Fanuc KAREL source: kt00240.KL

PROGRAM KT00240
%STACKSIZE=65535
%PRIORITY=65535
%NOLOCKGROUP
VAR
I1 : INTEGER
H2 : ARRAY[2] OF SHORT
OUT : INTEGER
BEGIN
I1=2
H2[1]=3
-- UNRESOLVED_PC line 10 opcodes [21 22 9D 33 B3 47 23] marker_code=35
END KT00240
